// TIA Portal V20 export
TYPE "T2_UDT_Hijo"
// Prueba IA 2: UDT hijo
   STRUCT
      Valor : Int;   // Valor
      Texto : String[10];   // Texto
   END_STRUCT;
END_TYPE
